// Builds the JSON payloads the PLC publishes. Each Write method leaves one complete document in
// the payload buffer and returns FALSE if it did not fit.
FUNCTION_BLOCK AlarmJsonWriter
VAR
    _Writer  : FB_JsonSaxWriter;
    _Payload : STRING(GVL_Mqtt.MaxPayloadLength);
    _Length  : UDINT;
END_VAR

METHOD PRIVATE AddAlarmMembers
// Every field of one alarm. raisedFileTime is a string: the value is too large for a JavaScript number.
VAR_IN_OUT CONSTANT
    Alarm : ST_PlcAlarm;
END_VAR
VAR
    Key            : STRING(127);
    EventClass     : STRING(80);
    Raised         : STRING(30);
    RaisedFileTime : STRING(24);
    Severity       : STRING(15);
    SeverityLevel  : DINT;
END_VAR
Key := F_AlarmKey(Alarm := Alarm);
EventClass := F_ToLCase(GUID_TO_STRING(Alarm.Entry.uuidEventClass));
Raised := F_FileTimeToIso(FileTime := Alarm.TimeRaised);
RaisedFileTime := ULINT_TO_STRING(Alarm.TimeRaised);

CASE Alarm.Entry.eSeverity OF
    TcEventSeverity.Verbose:
        Severity := 'Verbose';
        SeverityLevel := 0;
    TcEventSeverity.Info:
        Severity := 'Info';
        SeverityLevel := 1;
    TcEventSeverity.Warning:
        Severity := 'Warning';
        SeverityLevel := 2;
    TcEventSeverity.Error:
        Severity := 'Error';
        SeverityLevel := 3;
    TcEventSeverity.Critical:
        Severity := 'Critical';
        SeverityLevel := 4;
ELSE
    Severity := 'Unknown';
    SeverityLevel := -1;
END_CASE

_Writer.AddKey('key');
_Writer.AddString(Key);
_Writer.AddKey('eventClass');
_Writer.AddString(EventClass);
_Writer.AddKey('eventId');
_Writer.AddUdint(Alarm.Entry.nEventId);
_Writer.AddKey('severity');
_Writer.AddString(Severity);
_Writer.AddKey('severityLevel');
_Writer.AddDint(SeverityLevel);
_Writer.AddKey('source');
_Writer.AddString(Alarm.SourceName);
_Writer.AddKey('raised');
_Writer.AddString(Raised);
_Writer.AddKey('raisedFileTime');
_Writer.AddString(RaisedFileTime);
_Writer.AddKey('confirmed');
_Writer.AddBool(Alarm.IsConfirmed);
_Writer.AddKey('textAvailable');
_Writer.AddBool(Alarm.TextAvailable);
_Writer.AddKey('text');
_Writer.AddString(Alarm.Text);
END_METHOD

METHOD PRIVATE AddEnvelope
VAR_IN_OUT CONSTANT
    Envelope : ST_MqttEnvelope;
END_VAR
_Writer.AddKey('thing');
_Writer.AddString(Envelope.Thing);
_Writer.AddKey('session');
_Writer.AddString(Envelope.Session);
_Writer.AddKey('sequence');
_Writer.AddUdint(Envelope.Sequence);
_Writer.AddKey('timestamp');
_Writer.AddString(Envelope.Timestamp);
_Writer.AddKey('mode');
_Writer.AddString(Envelope.Mode);
IF LEN(Envelope.Reason) > 0 THEN
    _Writer.AddKey('reason');
    _Writer.AddString(Envelope.Reason);
END_IF
END_METHOD

METHOD PRIVATE Finish : BOOL
// Copies the document into the payload buffer, without the terminating null byte.
VAR
    Copied : UDINT;
END_VAR
Copied := _Writer.CopyDocument(pDoc := _Payload, nDoc := SIZEOF(_Payload));
_Writer.ResetDocument();
IF Copied > 1 THEN
    _Length := Copied - 1;
    Finish := TRUE;
ELSE
    _Length := 0;
    Finish := FALSE; // did not fit
END_IF
END_METHOD

PROPERTY PayloadAddress : PVOID
GET
PayloadAddress := ADR(_Payload);
END_GET
END_PROPERTY

PROPERTY PayloadLength : UDINT
GET
PayloadLength := _Length;
END_GET
END_PROPERTY

METHOD WriteAlarm : BOOL
// .../alarms/<key> in PerAlarm mode: one alarm.
VAR_IN_OUT CONSTANT
    Envelope : ST_MqttEnvelope;
    Alarm    : ST_PlcAlarm;
END_VAR
_Writer.ResetDocument();
_Writer.StartObject();
AddEnvelope(Envelope := Envelope);
AddAlarmMembers(Alarm := Alarm);
_Writer.EndObject();
WriteAlarm := Finish();
END_METHOD

METHOD WriteHeartbeat : BOOL
// .../heartbeat: the publisher is alive; how many alarms are raised.
VAR_IN_OUT CONSTANT
    Envelope : ST_MqttEnvelope;
END_VAR
VAR_INPUT
    Count    : UDINT;
    Overflow : BOOL;
END_VAR
_Writer.ResetDocument();
_Writer.StartObject();
AddEnvelope(Envelope := Envelope);
_Writer.AddKey('count');
_Writer.AddUdint(Count);
_Writer.AddKey('overflow');
_Writer.AddBool(Overflow);
_Writer.EndObject();
WriteHeartbeat := Finish();
END_METHOD

METHOD WriteIndex : BOOL
// .../alarms/index in PerAlarm mode: the keys of the current alarms.
VAR_IN_OUT CONSTANT
    Envelope : ST_MqttEnvelope;
    Keys     : ARRAY[0..GVL_EventLogging.MaxPlcAlarms - 1] OF STRING(127);
END_VAR
VAR_INPUT
    Count : UDINT;
END_VAR
VAR
    Row : DINT;
END_VAR
_Writer.ResetDocument();
_Writer.StartObject();
AddEnvelope(Envelope := Envelope);
_Writer.AddKey('count');
_Writer.AddUdint(Count);
_Writer.AddKey('keys');
_Writer.StartArray();
FOR Row := 0 TO UDINT_TO_DINT(Count) - 1 DO
    _Writer.AddString(Keys[Row]);
END_FOR
_Writer.EndArray();
_Writer.EndObject();
WriteIndex := Finish();
END_METHOD

METHOD WriteStatus : BOOL
// .../status: online or offline.
VAR_IN_OUT CONSTANT
    Envelope : ST_MqttEnvelope;
END_VAR
VAR_INPUT
    Online : BOOL;
END_VAR
_Writer.ResetDocument();
_Writer.StartObject();
AddEnvelope(Envelope := Envelope);
_Writer.AddKey('state');
IF Online THEN
    _Writer.AddString('online');
ELSE
    _Writer.AddString('offline');
END_IF
_Writer.EndObject();
WriteStatus := Finish();
END_METHOD

METHOD WriteTable : BOOL
// .../alarms in Table mode: every alarm in one document.
VAR_IN_OUT CONSTANT
    Envelope : ST_MqttEnvelope;
    Table    : ST_PlcAlarmTable;
END_VAR
VAR
    Row : DINT;
END_VAR
_Writer.ResetDocument();
_Writer.StartObject();
AddEnvelope(Envelope := Envelope);
_Writer.AddKey('count');
_Writer.AddUdint(Table.Count);
_Writer.AddKey('overflow');
_Writer.AddBool(Table.Overflow);
_Writer.AddKey('alarms');
_Writer.StartArray();
FOR Row := 0 TO UDINT_TO_DINT(Table.Count) - 1 DO
    _Writer.StartObject();
    AddAlarmMembers(Alarm := Table.Alarms[Row]);
    _Writer.EndObject();
END_FOR
_Writer.EndArray();
_Writer.EndObject();
WriteTable := Finish();
END_METHOD

END_FUNCTION_BLOCK

(* stored: Version 1.1.0.1, ProductVersion 3.1.4026.21
   POU AlarmJsonWriter: Id {c6761686-aefa-4076-9bbb-f5abb667b88e}, SpecialFunc None
   Method AddAlarmMembers: Id {d95fde15-4afb-4431-b998-e8d895482dc7}
   Method AddEnvelope: Id {8dfd5cf2-556f-437d-8e67-334d1a11a321}
   Method Finish: Id {b26ab69e-c499-4af9-a431-c719e84058d1}
   Property PayloadAddress: Id {91dedbe3-8f93-41d3-86ff-1654fea6e548}
   Get Get: Id {7bc3cfc2-8f3c-45a0-847b-2a68ff22c93e}
   Property PayloadLength: Id {c205bf7c-25e9-4182-a4f6-59897cae7979}
   Get Get: Id {8299018e-e0b9-4fa3-bb10-499c5a670930}
   Method WriteAlarm: Id {24f2973d-9511-44a7-aac6-08851f63ce68}
   Method WriteHeartbeat: Id {77303ce0-bfd7-4a4a-b76a-727c34eecfe1}
   Method WriteIndex: Id {bb548c19-596c-4888-b98a-1fce8742d058}
   Method WriteStatus: Id {95088f30-3cd8-4af8-bb9f-9f540f030bd2}
   Method WriteTable: Id {1dd3e349-5558-4c01-88da-d45840249b0d} *)
